Fanuc KAREL source: KA00218.KL

PROGRAM KA00218
%NOLOCKGROUP
VAR
  SRC: ARRAY[4] OF JOINTPOS
  DST: ARRAY[4] OF REAL
BEGIN
  DST = SRC
END KA00218
